(* IEC 61131-3 sources: rung/tests/conformance/cases, 12 files *)

(* ---- bits.st ---- *)
(* SPDX-License-Identifier: MIT *)
PROGRAM PRG_Bits
VAR CONSTANT
    cycles : UINT := 1;
END_VAR
VAR
    cycle : UINT;
    done : BOOL;
    b : BYTE := BYTE#16#81;
    w : WORD := WORD#16#8001;
    d : DWORD := DWORD#16#80000001;
    shift8 : UINT := 8;
    shift16 : UINT := 16;
    shift32 : UINT := 32;
    access : WORD := WORD#16#0008;
    (* SHL truncates a BYTE. *)
    r_byte_shl : BYTE;
    (* SHR shifts a BYTE logically. *)
    r_byte_shr : BYTE;
    (* SHL at the BYTE width. *)
    r_byte_width : BYTE;
    (* SHR beyond the BYTE width. *)
    r_byte_beyond : BYTE;
    (* SHL at the WORD width. *)
    r_word_width : WORD;
    (* SHR beyond the WORD width. *)
    r_word_beyond : WORD;
    (* SHL at the DWORD width exposes target-dependent shift counts. *)
    r_dword_width : DWORD;
    (* SHR beyond the DWORD width exposes target-dependent shift counts. *)
    r_dword_beyond : DWORD;
    (* WORD AND keeps only the low byte. *)
    r_and : WORD;
    (* WORD OR sets low bits. *)
    r_or : WORD;
    (* DWORD XOR complements all bits. *)
    r_xor : DWORD;
    (* DWORD NOT preserves unsigned width. *)
    r_not : DWORD;
    (* CODESYS bit access reads bit three. *)
    r_bit_read : BOOL;
    (* Bit assignment changes only the selected bit. *)
    r_bit_write : WORD;
END_VAR
IF NOT done THEN
    cycle := cycle + 1;
    r_byte_shl := SHL(b, 1);
    r_byte_shr := SHR(b, 1);
    r_byte_width := SHL(b, shift8);
    r_byte_beyond := SHR(b, shift8 + 1);
    r_word_width := SHL(w, shift16);
    r_word_beyond := SHR(w, shift16 + 1);
    r_dword_width := SHL(d, shift32);
    r_dword_beyond := SHR(d, shift32 + 1);
    r_and := w AND WORD#16#00FF;
    r_or := w OR WORD#16#00F0;
    r_xor := d XOR DWORD#16#FFFFFFFF;
    r_not := NOT d;
    r_bit_read := access.3;
    access.3 := FALSE;
    access.7 := TRUE;
    r_bit_write := access;
    done := cycle >= cycles;
END_IF
END_PROGRAM

(* ---- control.st ---- *)
(* SPDX-License-Identifier: MIT *)
PROGRAM PRG_Control
VAR CONSTANT
    cycles : UINT := 1;
END_VAR
VAR
    cycle : UINT;
    done : BOOL;
    selector : INT := 4;
    i : INT;
    total : INT;
    n : INT;
    (* CASE selects a range. *)
    r_case_range : INT;
    (* CASE selects an explicit list. *)
    r_case_list : INT;
    (* CASE falls back to ELSE. *)
    r_case_else : INT;
    (* FOR walks downward with a negative step. *)
    r_for_negative : INT;
    (* EXIT leaves FOR before its endpoint. *)
    r_for_exit : INT;
    (* CONTINUE skips the rest of a FOR iteration. *)
    r_for_continue : INT;
    (* WHILE tests its condition before each iteration. *)
    r_while : INT;
    (* REPEAT executes once when its condition starts true. *)
    r_repeat : INT;
    (* RETURN in an FC preserves the value already assigned. *)
    r_return_early : INT;
    (* The FC continues after a false RETURN condition. *)
    r_return_normal : INT;
END_VAR
IF NOT done THEN
    cycle := cycle + 1;
    CASE selector OF
        1..5: r_case_range := 11;
        ELSE r_case_range := 99;
    END_CASE
    CASE selector OF
        1, 4, 7: r_case_list := 22;
        ELSE r_case_list := 99;
    END_CASE
    CASE selector OF
        1, 2: r_case_else := 99;
        ELSE r_case_else := 33;
    END_CASE
    total := 0;
    FOR i := 5 TO -1 BY -2 DO
        total := total + i;
    END_FOR
    r_for_negative := total;
    total := 0;
    FOR i := 1 TO 10 DO
        IF i = 4 THEN EXIT; END_IF
        total := total + i;
    END_FOR
    r_for_exit := total;
    total := 0;
    FOR i := 1 TO 5 DO
        IF i = 3 THEN CONTINUE; END_IF
        total := total + i;
    END_FOR
    r_for_continue := total;
    n := 0;
    WHILE n < 4 DO
        n := n + 1;
    END_WHILE
    r_while := n;
    n := 5;
    REPEAT
        n := n + 1;
    UNTIL n >= 5
    END_REPEAT
    r_repeat := n;
    r_return_early := FC_ConformanceReturn(-3);
    r_return_normal := FC_ConformanceReturn(3);
    done := cycle >= cycles;
END_IF
END_PROGRAM

(* ---- conversions.st ---- *)
(* SPDX-License-Identifier: MIT *)
PROGRAM PRG_Conversions
VAR CONSTANT
    cycles : UINT := 1;
END_VAR
VAR
    cycle : UINT;
    done : BOOL;
    p_half : REAL := 0.5;
    p_one_half : REAL := 1.5;
    p_two_half : REAL := 2.5;
    n_half : REAL := -0.5;
    n_one_half : REAL := -1.5;
    n_two_half : REAL := -2.5;
    negative : REAL := -2.9;
    lp_half : LREAL := 2.5;
    ln_half : LREAL := -2.5;
    large : DINT := 16777217;
    integer : INT := -123;
    decimal_text : STRING := '-123';
    real_text : STRING := '12.5';
    typed_text : STRING := '16#FF';
    (* REAL_TO_INT at positive one half. *)
    r_half : INT;
    (* REAL_TO_INT at positive one and a half. *)
    r_one_half : INT;
    (* REAL_TO_INT at positive two and a half. *)
    r_two_half : INT;
    (* REAL_TO_INT at negative one half. *)
    r_neg_half : INT;
    (* REAL_TO_INT at negative one and a half. *)
    r_neg_one_half : INT;
    (* REAL_TO_INT at negative two and a half. *)
    r_neg_two_half : INT;
    (* LREAL_TO_DINT at a positive tie. *)
    r_lreal_half : DINT;
    (* LREAL_TO_DINT at a negative tie. *)
    r_lreal_neg_half : DINT;
    (* TRUNC discards a negative fractional part. *)
    r_trunc_neg : DINT;
    (* TRUNC at a positive rounding tie. *)
    r_trunc_tie : DINT;
    (* A negative INT converts to REAL. *)
    r_int_real : REAL;
    (* REAL loses the low bit beyond its 24-bit significand. *)
    r_real_precision : REAL;
    (* TRUE converts to one. *)
    r_bool_true : INT;
    (* FALSE converts to zero. *)
    r_bool_false : INT;
    (* Signed decimal STRING to INT. *)
    r_string_int : INT;
    (* Decimal STRING to REAL. *)
    r_string_real : REAL;
    (* Radix-prefixed STRING to UINT. *)
    r_string_hex : UINT;
    (* INT to signed decimal STRING. *)
    r_int_string : STRING;
    (* BOOL to STRING spelling. *)
    r_bool_string : STRING;
    (* REAL intermediate rounding is visible after cancellation. *)
    r_real_cancel : REAL;
END_VAR
IF NOT done THEN
    cycle := cycle + 1;
    r_half := REAL_TO_INT(p_half);
    r_one_half := REAL_TO_INT(p_one_half);
    r_two_half := REAL_TO_INT(p_two_half);
    r_neg_half := REAL_TO_INT(n_half);
    r_neg_one_half := REAL_TO_INT(n_one_half);
    r_neg_two_half := REAL_TO_INT(n_two_half);
    r_lreal_half := LREAL_TO_DINT(lp_half);
    r_lreal_neg_half := LREAL_TO_DINT(ln_half);
    r_trunc_neg := TRUNC(negative);
    r_trunc_tie := TRUNC(p_two_half);
    r_int_real := INT_TO_REAL(integer);
    r_real_precision := DINT_TO_REAL(large);
    r_bool_true := BOOL_TO_INT(TRUE);
    r_bool_false := BOOL_TO_INT(FALSE);
    r_string_int := STRING_TO_INT(decimal_text);
    r_string_real := STRING_TO_REAL(real_text);
    r_string_hex := STRING_TO_UINT(typed_text);
    r_int_string := INT_TO_STRING(integer);
    r_bool_string := BOOL_TO_STRING(TRUE);
    r_real_cancel := (DINT_TO_REAL(large) + REAL#1.0) - DINT_TO_REAL(large);
    done := cycle >= cycles;
END_IF
END_PROGRAM

(* ---- data.st ---- *)
(* SPDX-License-Identifier: MIT *)
PROGRAM PRG_Data
VAR CONSTANT
    cycles : UINT := 1;
END_VAR
VAR
    cycle : UINT;
    done : BOOL;
    a : ARRAY[-2..1] OF INT;
    grid : ARRAY[1..2, -1..1] OF INT;
    first : ST_ConformancePair;
    second : ST_ConformancePair;
    state : E_ConformanceState;
    i : INT;
    (* An array accepts a negative lower bound. *)
    r_array_low : INT;
    (* A FOR loop indexes every element across a non-zero lower bound. *)
    r_array_sum : INT;
    (* A multi-dimensional array preserves both lower bounds. *)
    r_grid : INT;
    (* Structure assignment copies members rather than aliasing. *)
    r_struct_number : INT;
    (* Structure assignment copies BOOL members. *)
    r_struct_flag : BOOL;
    (* An enumeration starts at its declared default. *)
    r_enum_default : INT;
    (* An enumeration member qualified by its type selects an explicit value. *)
    r_enum_typed : INT;
    (* CASE matches a qualified enumeration member. *)
    r_enum_case : INT;
END_VAR
IF NOT done THEN
    cycle := cycle + 1;
    a[-2] := 3;
    a[-1] := 5;
    a[0] := 7;
    a[1] := 11;
    r_array_low := a[-2];
    FOR i := -2 TO 1 DO
        r_array_sum := r_array_sum + a[i];
    END_FOR
    grid[1, -1] := 17;
    grid[2, 1] := 23;
    r_grid := grid[1, -1] + grid[2, 1];
    first.number := 12;
    first.flag := TRUE;
    second := first;
    first.number := 99;
    first.flag := FALSE;
    r_struct_number := second.number;
    r_struct_flag := second.flag;
    r_enum_default := state;
    state := E_ConformanceState.Running;
    r_enum_typed := state;
    CASE state OF
        E_ConformanceState.Running: r_enum_case := 42;
        ELSE r_enum_case := -1;
    END_CASE
    done := cycle >= cycles;
END_IF
END_PROGRAM

(* ---- int64.st ---- *)
(* SPDX-License-Identifier: MIT *)
PROGRAM PRG_Int64
VAR CONSTANT
    cycles : UINT := 1;
END_VAR
VAR
    cycle : UINT;
    done : BOOL;
    signed_high : LINT := LINT#4611686018427387904;
    unsigned_high : ULINT := ULINT#9223372036854775808;
    signed_min : LINT := LINT#-9223372036854775808;
    scratch : ULINT;
    (* A sum crossing the signed 64-bit boundary wraps. *)
    r_lint_overflow : LINT;
    (* Multiplication crossing the signed 64-bit boundary wraps. *)
    r_lint_mul : LINT;
    (* Negative LINT division preserves all 64 bits. *)
    r_lint_div : LINT;
    (* A sum crossing the unsigned 64-bit boundary wraps. *)
    r_ulint_overflow : ULINT;
    (* Multiplication crossing the unsigned 64-bit boundary wraps. *)
    r_ulint_mul : ULINT;
    (* Low bits of ULINT zero minus one; the full maximum is not a JavaScript integer. *)
    r_ulint_underflow_low : BYTE;
END_VAR
IF NOT done THEN
    cycle := cycle + 1;
    r_lint_overflow := signed_high + signed_high;
    r_lint_mul := signed_high * LINT#2;
    r_lint_div := signed_min / LINT#2;
    r_ulint_overflow := unsigned_high + unsigned_high;
    r_ulint_mul := unsigned_high * ULINT#2;
    scratch := ULINT#0;
    scratch := scratch - ULINT#1;
    r_ulint_underflow_low := ULINT_TO_BYTE(scratch);
    done := cycle >= cycles;
END_IF
END_PROGRAM

(* ---- rotates.st ---- *)
(* SPDX-License-Identifier: MIT *)
PROGRAM PRG_Rotates
VAR CONSTANT
    cycles : UINT := 1;
END_VAR
VAR
    cycle : UINT;
    done : BOOL;
    b : BYTE := BYTE#16#81;
    w : WORD := WORD#16#8001;
    d : DWORD := DWORD#16#80000001;
    width : UINT := 8;
    (* ROL carries the high BYTE bit into its low bit. *)
    r_byte_rol : BYTE;
    (* ROR carries the low BYTE bit into its high bit. *)
    r_byte_ror : BYTE;
    (* ROL by exactly the BYTE width. *)
    r_rol_width : BYTE;
    (* ROR beyond the BYTE width. *)
    r_ror_beyond : BYTE;
    (* ROL beyond the WORD width. *)
    r_word_rol : WORD;
    (* ROR beyond the DWORD width. *)
    r_dword_ror : DWORD;
END_VAR
IF NOT done THEN
    cycle := cycle + 1;
    r_byte_rol := ROL(b, 1);
    r_byte_ror := ROR(b, 1);
    r_rol_width := ROL(b, width);
    r_ror_beyond := ROR(b, width + 1);
    r_word_rol := ROL(w, 17);
    r_dword_ror := ROR(d, 33);
    done := cycle >= cycles;
END_IF
END_PROGRAM

(* ---- selection_math.st ---- *)
(* SPDX-License-Identifier: MIT *)
PROGRAM PRG_SelectionMath
VAR CONSTANT
    cycles : UINT := 1;
END_VAR
VAR
    cycle : UINT;
    done : BOOL;
    low : INT := -3;
    high : INT := 7;
    value : INT := 12;
    root : REAL := 2.0;
    base : LREAL := 2.0;
    (* Comparison of signed integers. *)
    r_less : BOOL;
    (* Equality of unequal values. *)
    r_equal : BOOL;
    (* Mixed REAL and LREAL comparison. *)
    r_real_cmp : BOOL;
    (* SEL false selects its first value. *)
    r_sel_false : INT;
    (* SEL true selects its second value. *)
    r_sel_true : INT;
    (* MUX zero selects the first value. *)
    r_mux_first : INT;
    (* MUX selects the last valid value. *)
    r_mux_last : INT;
    (* LIMIT clamps above the maximum. *)
    r_limit_high : INT;
    (* LIMIT clamps below the minimum. *)
    r_limit_low : INT;
    (* LIMIT preserves a value inside its bounds. *)
    r_limit_inside : INT;
    (* MIN accepts multiple operands. *)
    r_min : INT;
    (* MAX accepts multiple operands. *)
    r_max : INT;
    (* ABS of a negative INT. *)
    r_abs : INT;
    (* SQRT of a non-square REAL. *)
    r_sqrt : REAL;
    (* EXPT of an LREAL base. *)
    r_expt : LREAL;
END_VAR
IF NOT done THEN
    cycle := cycle + 1;
    r_less := low < high;
    r_equal := value = high;
    r_real_cmp := REAL#1.5 < LREAL#1.75;
    r_sel_false := SEL(FALSE, low, high);
    r_sel_true := SEL(TRUE, low, high);
    r_mux_first := MUX(0, low, high, value);
    r_mux_last := MUX(2, low, high, value);
    r_limit_high := LIMIT(low, value, high);
    r_limit_low := LIMIT(low, INT#-10, high);
    r_limit_inside := LIMIT(low, INT#2, high);
    r_min := MIN(value, low, high);
    r_max := MAX(value, low, high);
    r_abs := ABS(low);
    r_sqrt := SQRT(root);
    r_expt := EXPT(base, LREAL#3.0);
    done := cycle >= cycles;
END_IF
END_PROGRAM

(* ---- signed.st ---- *)
(* SPDX-License-Identifier: MIT *)
PROGRAM PRG_Signed
VAR CONSTANT
    cycles : UINT := 1;
END_VAR
VAR
    cycle : UINT;
    done : BOOL;
    sint_max : SINT := 127;
    sint_min : SINT := -128;
    int_max : INT := 32767;
    int_min : INT := -32768;
    dint_max : DINT := 2147483647;
    dint_min : DINT := -2147483648;
    dividend : INT := -7;
    divisor : INT := 3;
    small : SINT := 120;
    wider : DINT := 40000;
    (* SINT maximum plus one wraps on assignment. *)
    r_sint_overflow : SINT;
    (* SINT minimum minus one wraps on assignment. *)
    r_sint_underflow : SINT;
    (* SINT multiplication truncates to its destination width. *)
    r_sint_mul : SINT;
    (* INT maximum plus one wraps on assignment. *)
    r_int_overflow : INT;
    (* INT minimum minus one wraps on assignment. *)
    r_int_underflow : INT;
    (* INT multiplication truncates to its destination width. *)
    r_int_mul : INT;
    (* DINT maximum plus one wraps on assignment. *)
    r_dint_overflow : DINT;
    (* DINT minimum minus one wraps on assignment. *)
    r_dint_underflow : DINT;
    (* DINT multiplication truncates to its destination width. *)
    r_dint_mul : DINT;
    (* Integer division of a negative dividend truncates toward zero. *)
    r_div_negative : INT;
    (* A negative divisor reverses the quotient sign. *)
    r_div_negative_divisor : INT;
    (* MOD with a negative dividend. *)
    r_mod_negative : INT;
    (* MOD with a negative divisor. *)
    r_mod_negative_divisor : INT;
    (* Mixed SINT and DINT arithmetic widens before assignment. *)
    r_mixed_widen : DINT;
    (* An INT sum assigned to DINT exposes native intermediate width. *)
    r_intermediate : DINT;
END_VAR
IF NOT done THEN
    cycle := cycle + 1;
    r_sint_overflow := sint_max + SINT#1;
    r_sint_underflow := sint_min - SINT#1;
    r_sint_mul := sint_max * SINT#2;
    r_int_overflow := int_max + INT#1;
    r_int_underflow := int_min - INT#1;
    r_int_mul := int_max * INT#2;
    r_dint_overflow := dint_max + DINT#1;
    r_dint_underflow := dint_min - DINT#1;
    r_dint_mul := dint_max * DINT#2;
    r_div_negative := dividend / divisor;
    r_div_negative_divisor := dividend / -divisor;
    r_mod_negative := dividend MOD divisor;
    r_mod_negative_divisor := INT#7 MOD -divisor;
    r_mixed_widen := small + wider;
    r_intermediate := int_max + INT#1;
    done := cycle >= cycles;
END_IF
END_PROGRAM

(* ---- state.st ---- *)
(* SPDX-License-Identifier: MIT *)
PROGRAM PRG_State
VAR CONSTANT
    cycles : UINT := 8;
END_VAR
VAR
    cycle : UINT;
    done : BOOL;
    first : FB_ConformanceAccumulate;
    second : FB_ConformanceAccumulate;
    rising : R_TRIG;
    falling : F_TRIG;
    up : CTU;
    down : CTD;
    both : CTUD;
    set_latch : SR;
    reset_latch : RS;
    pulse : BOOL;
    (* An FB instance keeps its accumulator across cycles. *)
    r_fb_first : INT;
    (* Two instances of one FB keep independent state. *)
    r_fb_second : INT;
    (* R_TRIG fires once per rising edge. *)
    r_rising_count : INT;
    (* F_TRIG fires once per falling edge. *)
    r_falling_count : INT;
    (* F_TRIG on an initially false signal. *)
    r_falling_initial : BOOL;
    (* CTU reaches its preset after two edges. *)
    r_up_at_preset : WORD;
    (* CTU behavior on edges beyond its preset. *)
    r_up_after_preset : WORD;
    (* CTU Q at and beyond its preset. *)
    r_up_q : BOOL;
    (* CTD reaches zero from its loaded preset. *)
    r_down_zero : WORD;
    (* CTD behavior on an edge after reaching zero. *)
    r_down_after_zero : WORD;
    (* CTD Q after reaching zero. *)
    r_down_q : BOOL;
    (* CTUD handles simultaneous rising up and down edges. *)
    r_both_simultaneous : WORD;
    (* CTUD RESET and LOAD are asserted together. *)
    r_both_reset_load : WORD;
    (* CTUD upper output after reset. *)
    r_both_qu : BOOL;
    (* CTUD lower output after reset. *)
    r_both_qd : BOOL;
    (* SR is set dominant when both inputs are true. *)
    r_sr_both : BOOL;
    (* RS is reset dominant when both inputs are true. *)
    r_rs_both : BOOL;
    (* SR keeps its value after both inputs fall. *)
    r_sr_hold : BOOL;
    (* RS keeps its value after both inputs fall. *)
    r_rs_hold : BOOL;
END_VAR
IF NOT done THEN
    cycle := cycle + 1;
    pulse := (cycle MOD 2) = 0;
    first(increment := 1);
    second(increment := 3);
    r_fb_first := first.total;
    r_fb_second := second.total;
    rising(CLK := pulse);
    falling(CLK := pulse);
    IF rising.Q THEN r_rising_count := r_rising_count + 1; END_IF
    IF falling.Q THEN r_falling_count := r_falling_count + 1; END_IF
    IF cycle = 1 THEN r_falling_initial := falling.Q; END_IF
    up(CU := pulse, RESET := cycle = 1, PV := WORD#2);
    down(CD := pulse, LOAD := cycle = 1, PV := WORD#2);
    both(CU := pulse, CD := cycle = 4, RESET := cycle = 1 OR cycle = 8, LOAD := cycle = 8, PV := WORD#3);
    set_latch(SET1 := cycle = 2, RESET := cycle = 2);
    reset_latch(SET := cycle = 2, RESET1 := cycle = 2);
    IF cycle = 2 THEN
        r_sr_both := set_latch.Q1;
        r_rs_both := reset_latch.Q1;
    END_IF
    IF cycle = 3 THEN
        r_sr_hold := set_latch.Q1;
        r_rs_hold := reset_latch.Q1;
    END_IF
    IF cycle = 4 THEN
        r_up_at_preset := up.CV;
        r_down_zero := down.CV;
        r_both_simultaneous := both.CV;
    END_IF
    IF cycle = 6 THEN
        r_up_after_preset := up.CV;
        r_up_q := up.Q;
        r_down_after_zero := down.CV;
        r_down_q := down.Q;
    END_IF
    IF cycle = 8 THEN
        r_both_reset_load := both.CV;
        r_both_qu := both.QU;
        r_both_qd := both.QD;
    END_IF
    done := cycle >= cycles;
END_IF
END_PROGRAM

(* ---- strings.st ---- *)
(* SPDX-License-Identifier: MIT *)
PROGRAM PRG_Strings
VAR CONSTANT
    cycles : UINT := 1;
END_VAR
VAR
    cycle : UINT;
    done : BOOL;
    text : STRING := 'ABCDE';
    empty : STRING;
    (* LEN counts characters in a nonempty STRING. *)
    r_len : INT;
    (* LEN of an empty STRING. *)
    r_len_empty : INT;
    (* LEFT takes the first two characters. *)
    r_left : STRING;
    (* LEFT with zero length. *)
    r_left_zero : STRING;
    (* RIGHT takes the last two characters. *)
    r_right : STRING;
    (* RIGHT with a length beyond the input. *)
    r_right_long : STRING;
    (* MID uses a one-based start position. *)
    r_mid : STRING;
    (* MID at the last character. *)
    r_mid_last : STRING;
    (* MID starting beyond the input. *)
    r_mid_past : STRING;
    (* CONCAT appends a second STRING. *)
    r_concat : STRING;
    (* FIND returns a one-based position. *)
    r_find : INT;
    (* FIND returns zero when absent. *)
    r_find_missing : INT;
    (* FIND of an empty search STRING. *)
    r_find_empty : INT;
    (* INSERT follows its specified character. *)
    r_insert : STRING;
    (* INSERT at the last character. *)
    r_insert_end : STRING;
    (* DELETE removes two characters from position two. *)
    r_delete : STRING;
    (* DELETE at the last character. *)
    r_delete_last : STRING;
    (* REPLACE exchanges two characters at position two. *)
    r_replace : STRING;
    (* REPLACE grows a string at its last character. *)
    r_replace_last : STRING;
    (* INSERT at zero prepends text in CODESYS. *)
    r_insert_zero : STRING;
    (* DELETE starting beyond the input. *)
    r_delete_past : STRING;
    (* REPLACE at position zero exposes edge behavior. *)
    r_replace_zero : STRING;
END_VAR
IF NOT done THEN
    cycle := cycle + 1;
    r_len := LEN(text);
    r_len_empty := LEN(empty);
    r_left := LEFT(text, 2);
    r_left_zero := LEFT(text, 0);
    r_right := RIGHT(text, 2);
    r_right_long := RIGHT(text, 8);
    r_mid := MID(text, 2, 2);
    r_mid_last := MID(text, 1, 5);
    r_mid_past := MID(text, 2, 6);
    r_concat := CONCAT(text, '!');
    r_find := FIND(text, 'CD');
    r_find_missing := FIND(text, 'XY');
    r_find_empty := FIND(text, empty);
    r_insert := INSERT(text, 'xy', 2);
    r_insert_end := INSERT(text, 'xy', 5);
    r_delete := DELETE(text, 2, 2);
    r_delete_last := DELETE(text, 1, 5);
    r_replace := REPLACE(text, 'xy', 2, 2);
    r_replace_last := REPLACE(text, 'xy', 1, 5);
    r_insert_zero := INSERT(text, 'xy', 0);
    r_delete_past := DELETE(text, 2, 6);
    r_replace_zero := REPLACE(text, 'xy', 1, 0);
    done := cycle >= cycles;
END_IF
END_PROGRAM

(* ---- time.st ---- *)
(* SPDX-License-Identifier: MIT *)
PROGRAM PRG_Time
VAR CONSTANT
    cycles : UINT := 1;
END_VAR
VAR
    cycle : UINT;
    done : BOOL;
    one : TIME := T#1S;
    half : TIME := T#500MS;
    compound : TIME := T#1M2S3MS;
    (* TIME addition of seconds and milliseconds. *)
    r_add : TIME;
    (* TIME subtraction with a positive result. *)
    r_sub : TIME;
    (* Equivalent TIME literals compare equal. *)
    r_equal : BOOL;
    (* TIME ordering compares durations. *)
    r_less : BOOL;
    (* A compound TIME literal preserves milliseconds. *)
    r_compound : TIME;
    (* TIME to UDINT uses milliseconds. *)
    r_milliseconds : UDINT;
    (* MIN selects the shorter duration. *)
    r_min : TIME;
    (* LIMIT clamps a TIME duration. *)
    r_limit : TIME;
END_VAR
IF NOT done THEN
    cycle := cycle + 1;
    r_add := one + half;
    r_sub := one - half;
    r_equal := one + half = T#1500MS;
    r_less := half < one;
    r_compound := compound;
    r_milliseconds := TIME_TO_UDINT(compound);
    r_min := MIN(one, half);
    r_limit := LIMIT(half, T#2S, one);
    done := cycle >= cycles;
END_IF
END_PROGRAM

(* ---- unsigned.st ---- *)
(* SPDX-License-Identifier: MIT *)
PROGRAM PRG_Unsigned
VAR CONSTANT
    cycles : UINT := 1;
END_VAR
VAR
    cycle : UINT;
    done : BOOL;
    usint_max : USINT := 255;
    usint_zero : USINT;
    uint_max : UINT := 65535;
    uint_zero : UINT;
    udint_max : UDINT := 4294967295;
    udint_zero : UDINT;
    small : UINT := 65000;
    wide : UDINT := 100000;
    (* USINT maximum plus one wraps to zero. *)
    r_usint_overflow : USINT;
    (* USINT zero minus one wraps to the maximum. *)
    r_usint_underflow : USINT;
    (* USINT multiplication wraps at its width. *)
    r_usint_mul : USINT;
    (* UINT maximum plus one wraps to zero. *)
    r_uint_overflow : UINT;
    (* UINT zero minus one wraps to the maximum. *)
    r_uint_underflow : UINT;
    (* UINT multiplication wraps at its width. *)
    r_uint_mul : UINT;
    (* UDINT maximum plus one wraps to zero. *)
    r_udint_overflow : UDINT;
    (* UDINT zero minus one wraps to the maximum. *)
    r_udint_underflow : UDINT;
    (* UDINT multiplication wraps at its width. *)
    r_udint_mul : UDINT;
    (* UINT and UDINT arithmetic widens before assignment. *)
    r_mixed_widen : UDINT;
    (* A UINT sum assigned to UDINT exposes native intermediate width. *)
    r_intermediate : UDINT;
END_VAR
IF NOT done THEN
    cycle := cycle + 1;
    r_usint_overflow := usint_max + USINT#1;
    r_usint_underflow := usint_zero - USINT#1;
    r_usint_mul := usint_max * USINT#2;
    r_uint_overflow := uint_max + UINT#1;
    r_uint_underflow := uint_zero - UINT#1;
    r_uint_mul := uint_max * UINT#2;
    r_udint_overflow := udint_max + UDINT#1;
    r_udint_underflow := udint_zero - UDINT#1;
    r_udint_mul := udint_max * UDINT#2;
    r_mixed_widen := small + wide;
    r_intermediate := uint_max + UINT#1;
    done := cycle >= cycles;
END_IF
END_PROGRAM
